// TIA Portal V21 export
// export: Created 2026-10-14T03:09:03.0700016Z, ExportSetting WithDefaults, DisplayName Totally Integrated Automation Portal, DisplayVersion V21, DisplayName STEP 7 Professional, DisplayVersion V21, DisplayName STEP 7 Safety, DisplayVersion V21, DisplayName Tech WebApplication, DisplayVersion V21, DisplayName WinCC Basic/Comfort/Advanced, DisplayVersion V21, DisplayName WinCC Unified, DisplayVersion V21
TagTable "Filling"
  hmiStart : Bool  (HMI_Connection_1, 100 ms)
  hmiStop : Bool  (HMI_Connection_1, 100 ms)
  hmiReset : Bool  (HMI_Connection_1, 100 ms)
  tankLevel : Real  (HMI_Connection_1, 100 ms)
  tankTemperature : Real  (HMI_Connection_1, 100 ms)
  tankLevelMaxReached : Bool  (HMI_Connection_1, 100 ms)
  tankTempMax : Bool  (HMI_Connection_1, 100 ms)
  hmiNextBottle : Bool  (HMI_Connection_1, 100 ms)
  stateFillingTank : Bool  (HMI_Connection_1, 100 ms)
  stateHeatingTank : Bool  (HMI_Connection_1, 100 ms)
  stateFillingBottle : Bool  (HMI_Connection_1, 100 ms)
  stateShiftingBottle : Bool  (HMI_Connection_1, 100 ms)
  stateStop : Bool  (HMI_Connection_1, 100 ms)
  stateReset : Bool  (HMI_Connection_1, 100 ms)
  machineState : Int  (HMI_Connection_1, 100 ms)
  tankLevelMax : Real  (HMI_Connection_1, 100 ms)
  stateRunning : Bool  (HMI_Connection_1, 100 ms)
  bottleID : String  (HMI_Connection_1, 100 ms)
  bottlesProduced : UDInt  (HMI_Connection_1, 100 ms)
  bootleNumberFaulty : UDInt  (HMI_Connection_1, 100 ms)
  bottleLevel : Real  (HMI_Connection_1, 100 ms)
  HMI_bottleLevel1 : Real  (1 s)
  HMI_bottleLevel2 : Real  (1 s)
  HMI_bottleLevel3 : Real  (1 s)
  HMI_bottleLevel : Real  (HMI_Connection_1, 100 ms)
  HMI_doShift : Bool  (HMI_Connection_1, 100 ms)
    on ChangeValue: Conveyor()
  qrCode : String  (HMI_Connection_1, 100 ms)
  bottleFaulty : Bool  (HMI_Connection_1, 100 ms)
  qrCodeReceived : Bool  (HMI_Connection_1, 100 ms)
    on ChangeValue: HandleQrCode()
  tempInvisibleObject : Bool  (1 s, start 0)
  HMI_bottleInfo1 : Bool  (1 s)
  HMI_bottleInfo2 : Bool  (1 s)
  HMI_bottleInfo3 : Bool  (1 s)
  HMI_bottleInfo4 : Bool  (1 s)
  HMI_bottleInfoActive : Bool  (1 s)
  energyFillingTank : Real  (HMI_Connection_1, 100 ms)
  energyWaterFillingTank : Real  (HMI_Connection_1, 100 ms)
  energyHeatingTank : Real  (HMI_Connection_1, 100 ms)
  energyFillingBottles : Real  (HMI_Connection_1, 100 ms)
  tankPressure : Real  (HMI_Connection_1, 100 ms)
  stateError : Bool  (HMI_Connection_1, 100 ms)
  hmiError : Bool  (HMI_Connection_1, 100 ms)
  alarmIncoming : Bool  (HMI_Connection_1, 100 ms)
  batchID : UDInt  (HMI_Connection_1, 100 ms)
  energyGas : Real  (HMI_Connection_1, 100 ms)
